(* IEC 61131-3 sources: programs/VI-54/VI-54_20171205/VI-54_20171205/Stations/PLC_VI54/VI-54_171014/Class/SdiasSafetyBase, 1 file *)

(* ---- SdiasSafetyBase.st ---- *)
#include "..\..\Class\SdiasSafetyManager\SdiasSafetyManager.h"
#include "..\..\Class\SafetyBase\SafetyBase.h"
#include "..\..\Class\SdiasManager\SdiasManager.h"

(*!
<Class
	Name               = "SdiasSafetyBase"
	Revision           = "1.7"
	RealtimeTask       = "false"
	CyclicTask         = "false"
	BackgroundTask     = "false"
	Sigmatek           = "true"
	OSInterface        = "false"
	HighPriority       = "false"
	Automatic          = "false"
	UpdateMode         = "Prescan"
	IconPath           = ".\Class\Tool.ico"
	SharedCommandTable = "true"
	Objectsize         = "(586,120)">
	<Channels>
		<Server Name="CallCommand" Visualized="false" Initialize="false" WriteProtected="true" Retentive="false"/>
		<Server Name="ClassState" Visualized="true" Initialize="false" WriteProtected="true" Retentive="false"/>
		<Server Name="DeviceID" Visualized="true" Initialize="false" WriteProtected="true" Retentive="false" Comment="id of the detected device at this place"/>
		<Server Name="QuitComError" Visualized="true" Initialize="false" WriteProtected="false" Retentive="false" Comment="Write to this server to quit errors on safety cpu. &#13;&#10;It has the same function as QuitComError server on safety cpu.&#13;&#10;&#13;&#10;Server shows actual quit-state&#13;&#10;  2..busy with quitting general errors (safety dll version 6 or higher required)&#13;&#10;  1..busy with quitting communication error&#13;&#10;  0..ready&#13;&#10; -1..error at creating a new safety state&#13;&#10; -2..failed to disable user prompt for quit error&#13;&#10; -3..failed to select module via safety number&#13;&#10; -4..error at establishing connection to module (safety designer must not be online at the same time!)&#13;&#10; -5..failed to send the quit error command to the module&#13;&#10; -6..failed to delete the created safety state"/>
		<Server Name="RetryCounteruC1" Visualized="true" Initialize="false" WriteProtected="true" Retentive="false" Comment="Shows the amount of retry counters of microprocessor 1.&#13;&#10;-1 ... Retrycounter read out is not supported by this firmware version."/>
		<Server Name="RetryCounteruC2" Visualized="true" Initialize="false" WriteProtected="true" Retentive="false" Comment="Shows the amount of retry counters of microprocessor 2.&#13;&#10;-1 ... Retrycounter read out is not supported by this firmware version."/>
		<Server Name="SafetyNumber" Visualized="true" Initialize="false" WriteProtected="true" Retentive="false" Comment="This server shows the unique safety number of the hardware module"/>
		<Server Name="SerialNo" Class="String" Visualized="false" Initialize="false" WriteProtected="true" Retentive="false" Comment="This server shows the serial number of the hardware module."/>
		<Client Name="InputsNeeded" Required="true" Internal="false"/>
		<Client Name="OutputsNeeded" Required="true" Internal="false"/>
		<Client Name="Place" Required="true" Internal="false" Comment="place at SDIAS Safety bus (0..15)"/>
		<Client Name="Required" Required="false" Internal="false" DefValue="1" Comment="0 = module is not required&#13;&#10;1 = module is required (CPU will crash if module is missing)"/>
		<Client Name="SdiasSafetyIn" Required="true" Internal="false" Comment="This client must be connected to a SdiasSafetyOut Server of a SCP011 class"/>
		<Client Name="SerialNoStr" Required="true" Internal="true"/>
		<Client Name="SetDeviceID" Required="true" Internal="false"/>
	</Channels>
	<Dependencies>
		<Files>
			<File Path=".\Class\SdiasSafetyManager\SdiasSafetyManager.h" Include="true"/>
			<File Path=".\Class\SafetyBase\SafetyBase.h" Include="true"/>
			<File Path=".\Class\SdiasManager\SdiasManager.h" Include="true"/>
		</Files>
	</Dependencies>
	<RevDoku>
		<Owner Company="Sigmatek" Author="RamAnd"/>
		<Dokumentation Revision="1.7" Date="24.10.2016" Author="ZoePat" Company="Sigmatek" Description="Removed visualised-flag of server &quot;SerialNo&quot;, because the Server can not be used in the LSE. In excange the object of this class must be set to visualized in the derivations, to be able to visualize the embedded string object &quot;SerialNoStr&quot;."/>
		<Dokumentation Revision="1.6" Date="21.10.2014" Author="RamAnd" Company="Sigmatek" Description="Set Server QuitComError to visualized so it can be used in visualisation."/>
		<Dokumentation Revision="1.5" Date="31.10.2014" Author="lanste" Company="Sigmatek" Description="Added support to let derived classes react if the Hardware is not online."/>
		<Dokumentation Revision="1.4" Date="31.07.2014" Author="PieSte" Company="Sigmatek" Description="Added QuitComError server to quit errors on safety cpu."/>
		<Dokumentation Revision="1.3" Date="24.04.2014" Author="RamAnd" Company="Sigmatek" Description="Clear module info at the servers if a disconnect event occurs."/>
		<Dokumentation Revision="1.2" Date="22.04.2014" Author="EisMic" Company="Sigmatek" Description="Added new newinst command for safety retry counter."/>
		<Dokumentation Revision="1.1" Date="28.03.2014" Author="EisMic" Company="Sigmatek" Description="Added command in NewInst method of ClassState Server. Added servers RetryCounteruC1 and RetryCounteruC2."/>
		<Dokumentation Revision="1.0" Date="21.01.2014" Author="RamAnd" Company="Sigmatek" Description="First library version"/>
	</RevDoku>
	<Network Name="SdiasSafetyBase">
		<!-- List of Components in this network -->
		<Components>
			<Object
				Name       = "SerialNoStr"
				Class      = "String"
				Position   = "(240,300)"
				Visualized = "true">
				<Channels>
					<Server Name="Data"/>
					<Client Name="SingleRealloc" Value="1"/>
				</Channels>
			</Object>
		</Components>
		<Comments>
		</Comments>
		<!-- List of Connections in this network -->
		<Connections>
			<Connection Source="this.SerialNoStr" Destination="SerialNoStr.Data"/>
			<Connection Source="this.SerialNo" Destination="SerialNoStr.Data" Vertices="(728,330),(556,390),"/>
		</Connections>
		<!-- Headerfiles -->
		<Options>
		</Options>
	</Network>
</Class>
*)
SdiasSafetyBase : CLASS
  //Servers:
	ClassState 	: SvrChCmd_t_e_VaranErrors;
	DeviceID 	: SvrCh_UDINT;
	SerialNo 	: SvrChCmd_UDINT;
	SafetyNumber 	: SvrCh_HDINT;
	RetryCounteruC1 	: SvrCh_DINT;
	RetryCounteruC2 	: SvrCh_DINT;
	CallCommand 	: SvrChCmd_DINT;
	QuitComError 	: SvrCh_DINT;
  //Clients:
	SdiasSafetyIn 	: CltChCmd_DINT;
	Place 	: CltCh_UDINT;
	Required 	: CltCh_DINT;
	SetDeviceID 	: CltCh_DINT;
	InputsNeeded 	: CltCh_UDINT;
	OutputsNeeded 	: CltCh_UDINT;
	SerialNoStr 	: CltChCmd_String;
  //Variables:
		us_FirstScan 	: DINT;
		IOStates : BDINT
		[
		];

		UnsafeOutputStates : BDINT
		[
		];

		us_oldRetryCounteruc1 	: USINT;			//! <Variable Comment="Marker for old retry counter from microprocessor 1." Name="us_oldRetryCounteruc1"/>
		us_oldRetryCounteruc2 	: USINT;			//! <Variable Comment="Marker for old retry counter from microprocessor 2." Name="us_oldRetryCounteruc2"/>
  //Functions:

	FUNCTION SdiasSafetyBase
		VAR_OUTPUT
			ret_code 	: ConfStates;
		END_VAR;
				//! <Function Comment="Called when class state was set to _NoHardware &#13;&#10;No Implementation Overload in derived classes if needed " Name="SetClassStateError"/>
	FUNCTION VIRTUAL SetClassStateError;

	FUNCTION VIRTUAL GLOBAL Init;

	FUNCTION VIRTUAL GLOBAL RtWork
		VAR_INPUT
			EAX 	: UDINT;
		END_VAR
		VAR_OUTPUT
			state (EAX) 	: UDINT;
		END_VAR;

	FUNCTION VIRTUAL GLOBAL ClassState::NewInst
		VAR_INPUT
			pPara 	: ^CmdStruct;
			pResult 	: ^results;
		END_VAR
		VAR_OUTPUT
			ret_code 	: iprStates;
		END_VAR;

	FUNCTION VIRTUAL GLOBAL SerialNo::Read
		VAR_OUTPUT
			output (EAX) 	: UDINT;
		END_VAR;

	FUNCTION VIRTUAL GLOBAL SerialNo::Write
		VAR_INPUT
			input (EAX) 	: UDINT;
		END_VAR
		VAR_OUTPUT
			result (EAX) 	: UDINT;
		END_VAR;

	FUNCTION VIRTUAL GLOBAL CallCommand::NewInst
		VAR_INPUT
			pPara 	: ^CmdStruct;
			pResult 	: ^results;
		END_VAR
		VAR_OUTPUT
			ret_code 	: iprStates;
		END_VAR;

	FUNCTION VIRTUAL GLOBAL QuitComError::Write
		VAR_INPUT
			input (EAX) 	: DINT;
		END_VAR
		VAR_OUTPUT
			result (EAX) 	: DINT;
		END_VAR;
  //Tables:
	FUNCTION @STD
		VAR_OUTPUT
			ret_code	: CONFSTATES;
		END_VAR;
	FUNCTION GLOBAL TAB @CT_;
END_CLASS;

#pragma using String

FUNCTION VIRTUAL GLOBAL SdiasSafetyBase::Init
	VAR
		MyPara 	 : CmdStruct;
		MyResult : Results;
	END_VAR

#ifdef DEACTIVATED_LSL
  IF Place.Read() = DEACTIVATED_LSL THEN
    ClassState := _NoHardware;
    return;
  END_IF;
#endif

  us_FirstScan += 1;

  if us_FirstScan = 1 then

    Place         := Place.Read();
    Required    := required.Read();
    SetDeviceID := SetDeviceID.Read();

    MyPara.uiCmd := SDIAS_SAFETY_LOGIN;
    MyPara.aPara[0] := this$DINT;
    MyPara.aPara[1] := Place$DINT;
    MyPara.aPara[2] := SetDeviceID$USINT;
    MyPara.aPara[3] := Required;
    MyPara.aPara[4] := InputsNeeded$USINT;
    MyPara.aPara[5] := OutputsNeeded$USINT;
    MyPara.aPara[6] := (#IOStates)$DINT;
    MyPara.aPara[7] := (#UnsafeOutputStates)$DINT;

    if SdiasSafetyIn.NewInst(#MyPara, #MyResult) <> READY then
      TRACE("(SdiasSafetyBase::Init) Failed to login to SdiasSafetyManager!");
    end_if;
  end_if;

END_FUNCTION

FUNCTION SdiasSafetyBase::SdiasSafetyBase
	VAR_OUTPUT
		ret_code 	: ConfStates;
	END_VAR

  ClassState := _NotInitialized;

	ret_code := C_OK;

END_FUNCTION

FUNCTION VIRTUAL GLOBAL SdiasSafetyBase::RtWork
	VAR_INPUT
		EAX 	: UDINT;
	END_VAR
	VAR_OUTPUT
		state (EAX) 	: UDINT;
	END_VAR

  // overload this method to refresh the safe in- and outputs

	state := READY;

END_FUNCTION

FUNCTION VIRTUAL GLOBAL SdiasSafetyBase::ClassState::NewInst
	VAR_INPUT
		pPara 	: ^CmdStruct;
		pResult 	: ^Results;
	END_VAR
	VAR_OUTPUT
		ret_code 	: IprStates;
	END_VAR
  VAR
  	pSerNoStr : ^CHAR;
  END_VAR

	ret_code := READY;

	CASE pPara^.uiCmd OF
//**********************************************************************************************************************************************************
		SDIAS_SET_CLASS_STATE:

      // Only set "_ModuleFoundButManagerIsOff" if state = _ClassOk so that errorstates do not get overwriten
      if ( (pPara^.aPara[0]$t_e_VaranErrors = _ModuleFoundButManagerIsOff) &
           (ClassState <> _ClassOk) )  then
        return;
      end_if;

      ClassState := pPara^.aPara[0]$t_e_VaranErrors;
      DeviceID   := pPara^.aPara[1]$UDINT;

      // if the module has been disconnected => also delete the other infos about it
      if (ClassState = _NoHardware) then
        SerialNoStr.Clear();
        SafetyNumber := 0;

        // if we support retry counters => also reset them
        if RetryCounteruC1 <> -1 then
          RetryCounteruC1 := RetryCounteruC2 := 0;
          us_oldRetryCounteruc1 := us_oldRetryCounteruc2 := 0;
        end_if;

      end_if;

      if (ClassState <> _ClassOk) then
        // Let derived classes update their servers
        SetClassStateError();
      end_if;

//**********************************************************************************************************************************************************
    SDIAS_SET_NUMBERS:
      SafetyNumber := pPara^.aPara[0]$HDINT;
      pSerNoStr    := pPara^.aPara[1]$^CHAR;
      SerialNoStr.WriteDataOff(udLen:=_strlen(src:=pSerNoStr), udOff:=0, pData:=pSerNoStr);

//**********************************************************************************************************************************************************
    SDIAS_SET_RETRY_COUNTER:
    //Only Write if Retry counter has changed
    if pPara^.aPara[0] <> us_oldRetryCounteruc1 then
      //Add new amount and substract the old one
      RetryCounteruC1 += to_usint(pPara^.aPara[0] - us_oldRetryCounteruc1);
      us_oldRetryCounteruc1 := pPara^.aPara[0]$USINT;

    end_if;

    //Only Write if Retry counter has changed
    if pPara^.aPara[1] <> us_oldRetryCounteruc2 then
      //Add new amount and substract the old one
      RetryCounteruC2 += to_usint(pPara^.aPara[1] - us_oldRetryCounteruc2);
      us_oldRetryCounteruc2 := pPara^.aPara[1]$USINT;

    end_if;

//**********************************************************************************************************************************************************
    SDIAS_RETRY_COUNTER_NOT_AVAILABLE:
      RetryCounteruC1 := -1;
      RetryCounteruC2 := -1;

//**********************************************************************************************************************************************************
	  SDIAS_SET_ASY_STATE:
      QuitComError := pPara^.aPara[0]$^t_AsyRefresh^.QuitComError;

//**********************************************************************************************************************************************************
  END_CASE;

END_FUNCTION

FUNCTION VIRTUAL GLOBAL SdiasSafetyBase::CallCommand::NewInst
	VAR_INPUT
		pPara 	: ^CmdStruct;
		pResult 	: ^Results;
	END_VAR
	VAR_OUTPUT
		ret_code 	: IprStates;
	END_VAR

	ret_code := ERROR;

	CASE pPara^.uiCmd OF
//**********************************************************************************************************************************************************
    // forward commands from clients to manager
    SDIAS_CMD_ADD_RD_ACCESS,
    SDIAS_CMD_ADD_WR_ACCESS,
    SDIAS_CMD_SDO_SEND_REQUEST,
    SDIAS_CMD_CHANGE_LED_STATE,
    SDIAS_CMD_DA_RD_ACCESS,
    SDIAS_CMD_DA_WR_ACCESS,
    SDIAS_CMD_REQUIRED_ERROR,
    SDIAS_CMD_INIT_STATE_LOGIN,
    SDIAS_CMD_GET_HW_PATH,
    SDIAS_CMD_INSTALL_CYCLIC_TASK:
      ret_code := SdiasSafetyIn.NewInst(pPara, pResult);
//**********************************************************************************************************************************************************
	END_CASE;

END_FUNCTION

FUNCTION VIRTUAL GLOBAL SdiasSafetyBase::SerialNo::Read
	VAR_OUTPUT
		output (EAX) 	: UDINT;
	END_VAR

	SerialNo := SerialNoStr.Data.Read();
	output := SerialNo;

END_FUNCTION

FUNCTION VIRTUAL GLOBAL SdiasSafetyBase::SerialNo::Write
	VAR_INPUT
		input (EAX) 	: UDINT;
	END_VAR
	VAR_OUTPUT
		result (EAX) 	: UDINT;
	END_VAR

	SerialNo := input;
	result := (SerialNoStr.Data.Write(SerialNo))$UDINT;

END_FUNCTION

FUNCTION VIRTUAL GLOBAL SdiasSafetyBase::QuitComError::Write
	VAR_INPUT
		input (EAX) 	: DINT;
	END_VAR
	VAR_OUTPUT
		result (EAX) 	: DINT;
	END_VAR
  VAR
		MyPara 	  : CmdStruct;
		MyResult	: results;
  END_VAR

  QuitComError := input;
  // tell the outer class
  MyPara.uiCmd    := SDIAS_SET_QUITCOMERROR_IO;
  MyPara.aPara[0] := QuitComError;
  result$UDINT    := SdiasSafetyIn.NewInst(#MyPara, #MyResult);

END_FUNCTION

FUNCTION VIRTUAL SdiasSafetyBase::SetClassStateError

  // Called when class state was set to _NoHardware
  // No Implementation Overload in derived classes if needed

END_FUNCTION
